(* PLC project g_packaging_filler_clean, Anonymous Benchmark Suite 1.0 *)
(* stored: creationDateTime 2026-07-09T00:00:00 *)

PROGRAM g_packaging_filler_clean
  VAR_INPUT
    bottle_present : BOOL;
    full : BOOL;
    start : BOOL;
    maint : BOOL;
  END_VAR
  VAR_OUTPUT
    fill_valve : BOOL;
    reject : BOOL;
  END_VAR

(* LD diagram, written out as Structured Text *)
fill_valve := NOT full AND bottle_present AND start;
reject := NOT bottle_present AND start;
END_PROGRAM

CONFIGURATION Config0
  RESOURCE Res0 ON PLC
    TASK tcyclic(INTERVAL := T#10ms, PRIORITY := 0);
    PROGRAM inst0 WITH tcyclic : g_packaging_filler_clean;
  END_RESOURCE
END_CONFIGURATION
